// TIA Portal V20 export
// export: Created 2026-10-19T18:07:39.3920336Z, ExportSetting WithDefaults, DisplayName Totally Integrated Automation Portal, DisplayVersion V20 Update 6, DisplayName TIA Portal Openness, DisplayVersion V20 Update 6, DisplayName TIA Portal Version Control Interface, DisplayVersion V20 Update 6, DisplayName SINAMICS Startdrive Advanced, DisplayVersion V20 SP1, DisplayName SINAMICS Startdrive G130, G150, S120, S150, SINAMICS MV, G220, S200, S210, DisplayVersion V20 SP1, DisplayName SINAMICS Startdrive G110M, G120, G120C, G120D, G120P, G115D, DisplayVersion V20 SP1, DisplayName STEP 7 Professional, DisplayVersion V20 Update 6, DisplayName STEP 7 Safety, DisplayVersion V20 Update 2, DisplayName WinCC Basic/Comfort/Advanced, DisplayVersion V20 Update 6, DisplayName WinCC Unified, DisplayVersion V20 Update 6
DATA_BLOCK "SICK_Lector"   // DB46
{ S7_Optimized_Access := 'TRUE' }
VERSION : 0.1
// stored: AutoNumber true, DBAccessibleFromOPCUA true, DBAccessibleFromWebserver true, IsOnlyStoredInLoadMemory false, IsRetainMemResEnabled false, IsWriteProtectedInAS false, MemoryReserve 100
   VAR
      Barcode_Result : String;
      HWInputIdent : HW_IO := 554;
      HWInputLength : USInt := 32;
      HWOutputIdent : HW_IO := 555;
      HWOutputLength : USInt := 32;
      CANId : USInt := 0;
      TOut : Time := T#10S;
      Req : Bool := FALSE;
      TriggerOn : Bool := FALSE;
      TriggerOff : Bool := FALSE;
      Matchcode : Bool := FALSE;
      SavePermanent : Bool := FALSE;
      ComTest : Bool := FALSE;
      FreeCommand : Bool := FALSE;
      Data : "ST_SICK_Lector_CLV6xx";
      RdDone { S7_SetPoint := 'True'} : Bool := FALSE;
      ReqDone : Bool := FALSE;
      ReqBusy : Bool := FALSE;
      Error : Bool := TRUE;
      Errorcode : DWord := 16#0000_0015;
   END_VAR
BEGIN
   Data.Matchcode.sName := '';
   Data.Matchcode.nCodeType := ' ';
   Data.Matchcode.iMinMaxLength := 0;
   Data.Matchcode.sContent := '';
   Data.FreeCommand.sCommand := '';
   Data.FreeCommand.sResult := '';
   Data.ReadingResult.iCounter := 0;
   Data.ReadingResult.iLength := 0;
   Data.ReadingResult.arrResult[1..200] := 16#00;
END_DATA_BLOCK
